(* IEC 61131-3 sources: 2026_Projet_YGO_ExcavatriceDragage/TOOLS/LINTER_ST/stubs, 3 files *)

(* ---- DEVICE_STATE.st ---- *)
(* Type standard CODESYS IoStandard pour le Linter ST *)
TYPE DEVICE_STATE :
(
    UNKNOWN             := 0,
    STOPPED             := 1,
    CONFIG_ERROR        := 2,
    BUS_ERROR           := 3,
    DISABLED            := 4,
    INITIALIZING        := 5,
    RESET_ORIGIN        := 6,
    RESET_COMMUNICATION := 7,
    RESET_APPLICATION   := 8,
    RUNNING             := 9,
    LOGGER_ERROR        := 10
);
END_TYPE

(* ---- GVL_Device_IO.st ---- *)
VAR_GLOBAL
    // === 📥 ENTRÉES MATÉRIELLES (HwReal) ===

    // Treuils M1 / M2
    M1_ContactorsReleased_DI     : BOOL;
    M1_ThermalOk_DI              : BOOL;
    M1_BrakeIsOpen_DI            : BOOL;
    M2_ContactorsReleased_DI     : BOOL;
    M2_ThermalOk_DI              : BOOL;
    M2_BrakeIsOpen_DI            : BOOL;
    M1M2_TopPositionFree_DI      : BOOL;
    M2_TensionedCable_DI         : BOOL;

    // Codeurs absolus
    COD1_PosValue                : DINT;
    COD1_Alarms                  : DWORD;
    COD1_Warnings                : DWORD;
    COD1_PresetTTrigCmd          : BOOL;
    COD1_CodeSeqTrigCmd          : BOOL;
    COD1_PresetValue             : DINT;
    COD1_CODEUR                  : FB_DeviceStub;

    COD2_PosValue                : DINT;
    COD2_Alarms                  : DWORD;
    COD2_Warnings                : DWORD;
    COD2_PresetTTrigCmd          : BOOL;
    COD2_CodeSeqTrigCmd          : BOOL;
    COD2_PresetValue             : DINT;
    COD2_CODEUR                  : FB_DeviceStub;

    // Translation M3 (AC600)
    M3_PosTremie_DI              : BOOL;
    M3_PosPV_DI                  : BOOL;
    M3_PosPVP2_DI                : BOOL;
    M3_PosP1_DI                  : BOOL;
    M3_PosMaintenance_DI         : BOOL;
    M3_BrakeIsOpen_DI            : BOOL;
    M3_ThermalOK_DI              : BOOL;
    M3_StatusWord                : WORD;
    M3_ActualFrequencyHz         : WORD;
    AC600_ECAT_Drive             : FB_DeviceStub;

    // Joystick Opérateur / CANopen
    JoyXRaw_ANA1                 : INT;
    JoyYRaw_ANA2                 : INT;
    JoyBtnRaw                    : WORD;
    CANbus                       : FB_DeviceStub;
    JOY1_JOYSTICK_MCB560_CO4201A : FB_DeviceStub;

    // Sécurités / Communs Machine
    PowerContactorEngaged_DI     : BOOL;
    EmergencyChainClosed_DI      : BOOL;
    PhaseRotationOk_DI           : BOOL;
    M1_M2_M3_BrakeThermalOk_DI   : BOOL;
    M1_M2_KoboldBottomTouch_DI   : BOOL;
    HydraulicThermalOk_DI        : BOOL;
    ConveyorInfeedReady_DI       : BOOL;
    TremieFull_OR_GateRaised_DI  : BOOL;

    // Modules d'E/S déportées
    Local_Digital_IO             : FB_DeviceStub;
    VH_0800END                   : FB_DeviceStub;
    VH_0808ETP                   : FB_DeviceStub;
    VH_0008ER                    : FB_DeviceStub;
    VH_0008ER_1                  : FB_DeviceStub;

    // === 📤 SORTIES MATÉRIELLES (PRG_06_Outputs) ===

    // Treuil M1 (Retenue)
    M1_RelayAscent_RQ            : BOOL;
    M1_RelayDescent_RQ           : BOOL;
    M1_SpeedContactor_1_DQ       : BOOL;
    M1_SpeedContactor_2_DQ       : BOOL;
    M1_SpeedContactor_3_DQ       : BOOL;
    M1_SpeedContactor_4_DQ       : BOOL;
    M1_BrakeRelease_RQ           : BOOL;

    // Treuil M2 (Benne)
    M2_RelayAscent_Close_RQ      : BOOL;
    M2_RelayDescent_Open_RQ      : BOOL;
    M2_SpeedContactor_1_DQ       : BOOL;
    M2_SpeedContactor_2_DQ       : BOOL;
    M2_SpeedContactor_3_DQ       : BOOL;
    M2_SpeedContactor_4_DQ       : BOOL;
    M2_BrakeRelease_RQ           : BOOL;

    // Translation M3
    M3_CommandWord               : WORD;
    M3_SetpointFrequencyHz       : WORD;
    M3_BrakeRelease_RQ           : BOOL;

    // Capteur fond Kobold
    M1_M2_KoboldMeasureEnable_RQ : BOOL;

    // Chaîne Arrêt d'Urgence / Puissance
    PowerKeepAlive_A_RQ          : BOOL;
    PowerKeepAlive_B_RQ          : BOOL;
    EmergencyArming_RQ           : BOOL;
END_VAR

(* ---- FB_DeviceStub.st ---- *)
FUNCTION_BLOCK FB_DeviceStub
VAR_INPUT
END_VAR
VAR_OUTPUT
END_VAR
METHOD GetDeviceState : DEVICE_STATE
    GetDeviceState := DEVICE_STATE.RUNNING;
END_METHOD
METHOD GetBusState : DEVICE_STATE
    GetBusState := DEVICE_STATE.RUNNING;
END_METHOD
END_FUNCTION_BLOCK
